(* IEC 61131-3 sources: PLC-IsaVODE/PLC-IsaVODE/samples/proofs, 4 files *)

(* ---- 1-water_tank.st ---- *)
PROGRAM WTT
    VAR_INPUT
        x1, x2, f1, f2 : REAL;
    END_VAR
    VAR_OUTPUT
        V1, V2, P : BOOL;
    END_VAR

    IF (x1 >= H1) THEN
        V1 := 0;            (* Close inlet valve V1 if tank1 at high level *)
    ELSE
        IF (x1 <= L1) THEN
            V1 := 1;        (* Open V1 if tank1 at low level *)
        END_IF;
    END_IF;
    IF (x2 <= L2) THEN
        P := 1; V2 := 1;    (* If tank2 low, start pump P and open outlet valve V2 *)
    END_IF;
    IF (x1 <= LL OR f2 <= FL OR x2 >= H2) THEN
        P := 0; V2 := 0;    (* Emergency stop pump P and close V2 on underflow/overflow *)
    END_IF;
END_PROGRAM

(* ---- 3-bohlender-artcile-reset-example-safe.st ---- *)
PROGRAM RESET_BOHLENDER
	VAR RETAIN
	    fs : bool := true;
		b : int := 0;
	END_VAR
	VAR
	    a : int := 0;
	END_VAR

    IF fs THEN
    	b := 2;
    	fs := false;
    END_IF;
    a := 1234 / b;
END_PROGRAM

(* ---- 3-bohlender-artcile-reset-example.st ---- *)
PROGRAM RESET_BOHLENDER
	VAR RETAIN
	    fs : bool := true;
	END_VAR
	VAR
	    a : int := 0;
		b : int := 0;
	END_VAR

    IF fs THEN
    	b := 2;
    	fs := false;
    END_IF;
    a := 1234 / b;
END_PROGRAM

(* ---- 4-calibrate.st ---- *)
PROGRAM CALIBRATE
	VAR_INPUT
		X        : REAL;
		CO       : BOOL;
		CS       : BOOL;
		Y_OFFSET : REAL;
		Y_SCALE  : REAL;
	END_VAR

	VAR_OUTPUT
		Y 		 : REAL;
	END_VAR

	VAR RETAIN
		OFFSET   : REAL;
		SCALE    : REAL := 1.0;
	END_VAR

	IF CO THEN
		OFFSET := Y_OFFSET - X;
	ELSIF CS THEN
		SCALE := Y_SCALE / (X + OFFSET);
	END_IF;
	Y := (X + OFFSET) * SCALE;

END_PROGRAM
